FUNCTION_BLOCK HANDWIRED_RUN (* Runs a program file exported by handwired-rs: the same operations in the same order on every input, refusing inputs outside its function's ranges, grids and types *)
  (* Description: SPDX-License-Identifier: MIT *)
  (* Version 0.1, 2026-11-19, handwired-rs, handwired-rs *)
  PACKAGE handwired;
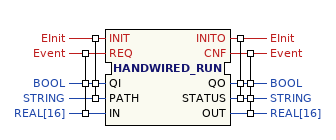
  EVENT_INPUT
    INIT : EInit WITH QI, PATH; (* QI = TRUE: read and check the program file at PATH; QI = FALSE: unload it *)
    REQ WITH QI, IN; (* Run the program on the first cells of IN *)
  END_EVENT
  EVENT_OUTPUT
    INITO : EInit WITH QO, STATUS; (* Loaded (QO = TRUE) or not, and why *)
    CNF WITH QO, STATUS, OUT; (* Ran (QO = TRUE, OUT written) or refused (QO = FALSE, OUT unchanged) *)
  END_EVENT
  VAR_INPUT
    QI : BOOL; (* Event input qualifier *)
    PATH : STRING; (* The program file (.hwc), relative to FORTE's working directory *)
    IN : ARRAY [0..15] OF REAL; (* Input cells; the program uses as many as it has inputs *)
  END_VAR
  VAR_OUTPUT
    QO : BOOL; (* Event output qualifier: FALSE when not loaded or refused *)
    STATUS : STRING; (* OK, the program's name and size after INIT, or why it was refused *)
    OUT : ARRAY [0..15] OF REAL; (* Output cells; the program writes as many as it has outputs *)
  END_VAR
END_FUNCTION_BLOCK
